TYPE e_DualChanal :(
	Wrong:=0,
	Close:=1,
	Open:=2);
END_TYPE

(* stored: Version 1.1.0.1, ProductVersion 3.1.4024.12
   DUT e_DualChanal: Id {c7c816e5-e291-49d4-9ac8-eeb98ef366ae} *)
